// TIA Portal V21 export
// export: Created 2026-10-23T20:42:29.8996432Z, ExportSetting WithDefaults, DisplayName Totally Integrated Automation Portal, DisplayVersion V21 Update 1, DisplayName SINAMICS Startdrive Advanced, DisplayVersion V21 HF2, DisplayName SINAMICS Startdrive G110M, G120, G120C, G120D, G120P, G115D, DisplayVersion V21 HF2, DisplayName SINAMICS Startdrive G130, G150, S120, S150, G200, G220, S200, S210, S220, Innomotics MVD, DisplayVersion V21 HF2, DisplayName STEP 7 Professional, DisplayVersion V21 Update 1, DisplayName STEP 7 Safety, DisplayVersion V21, DisplayName Tech WebApplication, DisplayVersion V21, DisplayName WinCC Basic/Comfort/Advanced, DisplayVersion V21 Update 1, DisplayName WinCC Unified, DisplayVersion V21 Update 1
FUNCTION "FC_IecOff" : Word   // FC4, SCL
TITLE = Implicit conversions, IEC check off
{ S7_Optimized_Access := 'TRUE' }
VERSION : 0.1
// Same body as FC_IecOn; this block has the IEC check switched off
// stored: AutoNumber true, IsIECCheckEnabled false, SetENOAutomatically false, UDAEnableTagReadback false
   VAR_INPUT
      InInt : Int;   // Integer input
      InWord : Word;   // Bit string input
      InDInt : DInt;   // Double integer input
   END_VAR
   VAR_OUTPUT
      OutInt : Int;   // Integer output
      OutSInt : SInt;   // Short integer output
      OutNarrow : Int;   // Narrowed double integer
   END_VAR
BEGIN

       // Implicit conversions between bit strings and integers, and narrowing conversions
       #OutInt := #InWord;
       #OutSInt := #InInt;
       #OutNarrow := #InDInt;
       #FC_IecOff := #InInt;
END_FUNCTION
